{region 'Documentation'}
(*!
<summary>Checks whether the ULINT value is inside the inclusive range.</summary>
<description>

Minimum &gt; Maximum reports Error during active evaluation; equal bounds are
valid.

</description>
*)
{endregion}
FUNCTION_BLOCK AssertInRange_ULInt EXTENDS AssertionBase
VAR_INPUT
    IN : ULINT; //! Actual value checked or observed by this Assertion.
    Minimum : ULINT; //! Inclusive lower bound of the comparison; for a range, must not exceed Maximum.
    Maximum : ULINT; //! Inclusive upper bound of the comparison; for a range, must not be below Minimum.
END_VAR

SUPER^();

{region 'Documentation'}
(*!
<summary>Check whether the ULINT value is inside the inclusive range.</summary>
*)
{endregion}
METHOD PROTECTED Assert
VAR
    Message : STRING(GVL_Constants.MessageLength);
    MinimumText : STRING(GVL_Constants.AssertionValueLength);
    MaximumText : STRING(GVL_Constants.AssertionValueLength);
    ActualText : STRING(GVL_Constants.AssertionValueLength);
END_VAR
IF NOT EvaluationActive THEN
    RETURN;
END_IF;

IF Result = E_Result.Error THEN
    RETURN;
END_IF;

IF Minimum > Maximum THEN
    MinimumText := ULINT_TO_STRING(Minimum);
    MaximumText := ULINT_TO_STRING(Maximum);
    Message := CONCAT('Assertion error: minimum exceeds maximum. Minimum = ',
        MinimumText);
    Message := CONCAT(Message, ', Maximum = ');
    Message := CONCAT(Message, MaximumText);
    Message := CONCAT(Message, '.');
    Error(Message := Message);
    RETURN;
END_IF;

IF Result = E_Result.Failed THEN
    RETURN;
END_IF;

IF (IN < Minimum) OR (IN > Maximum) THEN
    MinimumText := ULINT_TO_STRING(Minimum);
    MaximumText := ULINT_TO_STRING(Maximum);
    ActualText := ULINT_TO_STRING(IN);
    Message := CONCAT('Assertion failed: value is outside allowed range. Minimum = ',
        MinimumText);
    Message := CONCAT(Message, ', Maximum = ');
    Message := CONCAT(Message, MaximumText);
    Message := CONCAT(Message, ', Actual = ');
    Message := CONCAT(Message, ActualText);
    Message := CONCAT(Message, '.');
    Fail(Message := Message);
    RETURN;
END_IF;

Pass();
END_METHOD

END_FUNCTION_BLOCK

(* stored: Version 1.1.0.1
   POU AssertInRange_ULInt: Id {717bbeff-a017-4c5c-8dd5-dc334f429d77}, SpecialFunc None
   Folder Internal: Id {6379f793-58d7-42d1-873a-d46fd1ce93f7}
   Method Assert: Id {cd5eceea-0b2d-4073-8148-ee7815c47340} *)
